Universal Robots URScript: dual_arm_kitting_right.script

def right():
  # Generated by botrail (units: rad, m, s)
  # joints: right_shoulder_pan_joint, right_shoulder_lift_joint, right_elbow_joint, right_wrist_1_joint, right_wrist_2_joint, right_wrist_3_joint
  movej([0, -1.9, 1.8, -1.5, -1.57, 0], a=6.283185, v=3.141593, r=0)
  # step 1: right claim R1
  set_standard_digital_out(0, True)
  # step 2: right pick R1
  movej([-0.091113, -1.219699, 2.182763, -2.533862, -1.570796, -1.661909], a=6.283185, v=3.141593, r=0)
  movel([-0.091112, -0.960625, 2.202763, -2.812934, -1.570796, -1.661909], a=1.2, v=0.25, r=0)
  # step 3: right grasp R1
  # attach R1 (simulation grasp — drive the real gripper via a mapped output)
  # step 4: right wait bin R1
  while (get_standard_digital_in(0)):
    sync()
  end
  # step 5: right place R1
  movel([-0.091113, -1.219698, 2.182765, -2.533867, -1.570796, -1.661909], a=1.2, v=0.25, r=0)
  movej([0.479932, -1.735656, 2.440569, -2.275706, -1.570796, -1.090864], a=6.283185, v=3.141593, r=0)
  # step 6: right release R1
  # detach R1 (simulation release)
  set_standard_digital_out(0, False)
  # step 7: right clear R1
  movej([0, -1.9, 1.8, -1.5, -1.57, 0], a=6.283185, v=3.141593, r=0)
  # step 8: right claim R2
  set_standard_digital_out(0, True)
  # step 9: right pick R2
  movej([-0.070256, -0.98522, 1.769778, -2.355359, -1.570796, -1.641052], a=6.283185, v=3.141593, r=0)
  movel([-0.070255, -0.798708, 1.786383, -2.558465, -1.570796, -1.641052], a=1.2, v=0.25, r=0)
  # step 10: right grasp R2
  # attach R2 (simulation grasp — drive the real gripper via a mapped output)
  # step 11: right wait bin R2
  while (get_standard_digital_in(0)):
    sync()
  end
  # step 12: right place R2
  movel([-0.070259, -0.985224, 1.769811, -2.355403, -1.570795, -1.641055], a=1.2, v=0.25, r=0)
  movej([0.406587, -1.619605, 2.342258, -2.293448, -1.570796, -1.164209], a=6.283185, v=3.141593, r=0)
  # step 13: right release R2
  # detach R2 (simulation release)
  set_standard_digital_out(0, False)
  # step 14: right clear R2
  movej([0, -1.9, 1.8, -1.5, -1.57, 0], a=6.283185, v=3.141593, r=0)
  # step 15: right await handoff
  while (not get_standard_digital_in(1)):
    sync()
  end
  # step 16: right claim H
  set_standard_digital_out(0, True)
  # step 17: right pick H
  movej([0.284937, -0.990288, 1.768326, -2.348836, -1.570796, -1.285859], a=6.283185, v=3.141593, r=0)
  movel([0.284937, -0.804729, 1.786777, -2.552838, -1.570796, -1.285859], a=1.2, v=0.25, r=0)
  # step 18: right grasp H
  # attach L2 (simulation grasp — drive the real gripper via a mapped output)
  # step 19: right wait bin H
  while (get_standard_digital_in(0)):
    sync()
  end
  # step 20: right place H
  movel([0.284934, -0.990291, 1.768359, -2.34888, -1.570795, -1.285862], a=1.2, v=0.25, r=0)
  movej([0.54154, -1.512983, 2.234952, -2.292766, -1.570796, -1.029256], a=6.283185, v=3.141593, r=0)
  # step 21: right release H
  # detach L2 (simulation release)
  set_standard_digital_out(0, False)
  # step 22: right clear H
  movej([0, -1.9, 1.8, -1.5, -1.57, 0], a=6.283185, v=3.141593, r=0)
  # step 23: right cleared H
  set_standard_digital_out(1, True)
end
